(* IEC 61131-3 sources: 2026_Projet_YGO_ExcavatriceDragage/CODE_BACKUP/CODE_20260803_avant_ee4d08b/CODEURS, 7 files *)

(* ---- ST_Encoder_Calib.st ---- *)
(* ═══════════════════════════════════════════════════════════════
   🧲 ST_Encoder_Calib — Calibration & référence codeur (1 par treuil, RETAIN)
   ───────────────────────────────────────────────────────────────
   📄 Doc métier : DOC/AF_Partie-09_Fonction_Encoder_v2.1.md
                   DOC/AF_Partie-03_Contrats_Composants_v2.0.md
   🎛️ Une instance RETAIN par treuil (M1_EncoderCalib / M2_EncoderCalib).
   ═══════════════════════════════════════════════════════════════ *)

TYPE ST_Encoder_Calib :
STRUCT
    HomingRefRaw                  : UDINT;   // Valeur brute figée au dernier homing réussi
    LastKnownRawPos                : UDINT;   // Dernier point brut valide connu (§3.7, continu)
    RestartCoherenceTolerancePts    : UDINT := 1000;  // Tolérance redémarrage (~12% PointsPerRev 8192)
    Homed                          : BOOL;    // TRUE dès qu'un référencement a réussi
    HomingSuspect                  : BOOL;    // TRUE si incohérence détectée au redémarrage (§3.7)
END_STRUCT
END_TYPE

(* ---- FB_Encoder_Abs.st ---- *)
(* ═══════════════════════════════════════════════════════════════
   🧲 FB_Encoder_Abs — Acquisition codeur absolu (accès bus EtherCAT)
   ───────────────────────────────────────────────────────────────
   📄 Doc métier : DOC/AF_Partie-09_Fonction_Encoder_v2.1.md §3/§6
                   DOC/AF_Partie-03_Contrats_Composants_v2.0.md
   🎯 Accès bus EtherCAT, statut esclave, extraction positions brutes
      et séquence de Preset SDO (PresetTriggerCmd := 2).
   🧊 Principe « geler sur doute » (§6) : RawPos/AngleRaw/TurnCount
      conservent leur dernière valeur valide si EncoderAvailable = FALSE.
   ═══════════════════════════════════════════════════════════════ *)

// === DECLARATION (à coller dans la partie déclaration du POU FB_Encoder_Abs) ===

FUNCTION_BLOCK PUBLIC FB_Encoder_Abs
VAR_INPUT
    Enable              : BOOL;        // Standard
    Reset               : BOOL;        // Acquittement défaut (front)
    PowerContactorEngaged     : BOOL;        // Standard
    Mode                : E_Mode;      // Standard (contexte, pas encore exploité ce lot)
    RawPosIn            : UDINT;       // Brut EtherCAT (ex. COD1_PosValue, %ID)
    AlarmsIn            : UINT;        // Brut EtherCAT (ex. COD1_Alarms)
    WarningsIn          : UINT;        // Brut EtherCAT (ex. COD1_Warnings) — informatif seulement
    SlaveOperational    : BOOL;        // FB_Diag_Ethercat — esclave EtherCAT opérationnel
    PointsPerRev        : UDINT := 8192;  // Résolution codeur confirmée (Partie10 §3.3)
    PresetRequest       : BOOL;        // Front — piloté par FB_Encoder_Homing via PRG_02_Encoders
    PresetValue         : UDINT;       // Cible brute — piloté par FB_Encoder_Homing (stub 0 ce lot)
    PresetTimeout       : TIME := T#2s;
    PresetTolerancePts  : UDINT := 10; // Tolérance relecture post-preset
END_VAR
VAR_OUTPUT
    Ready               : BOOL;
    Busy                : BOOL;
    Done                : BOOL;
    Error               : BOOL;
    ErrorId             : WORD;        // bit0: "Défaut communication codeur" - alarme/bus codeur ; bit1: "Erreur référencement (timeout)" - preset refusé/timeout
    State               : E_State;
    StateAtError        : E_State;
    RawPos              : UDINT;       // Position brute — GELÉE si EncoderAvailable=FALSE
    EncoderAvailable    : BOOL;
    AngleRaw            : UINT;        // Informatif maintenance : RawPos MOD PointsPerRev
    TurnCount           : UDINT;       // Informatif maintenance : RawPos / PointsPerRev
    PresetAck           : BOOL;        // Pulse 1 cycle — écriture confirmée
    PresetNak           : BOOL;        // Pulse 1 cycle — écriture refusée/timeout
    PresetTriggerCmd    : WORD;        // → à câbler sur COD_PresettTrigCmd (RxPDO)
    CodeSeqTriggerCmd   : WORD;        // → à câbler sur COD_CodeSeqTrigCmd (RxPDO)
    PresetValueOut      : UDINT;       // → à câbler sur COD_PresetValue (RxPDO)
END_VAR
VAR
    ResetEdge           : R_TRIG;
    ErrorEdge           : R_TRIG;
    PresetReqEdge       : R_TRIG;
    PresetTimer         : TON;
    PresetSeqStep       : INT;         // 0=IDLE, 1=pulse CodeSeq, 2=pulse Trig, 3=attente confirmation
    RawDiff             : DINT;
    PresetTimerVisual   : TON;         // Timer pour laisser le temps de voir l'impulsion (1.5s)
END_VAR

// === IMPLEMENTATION (à coller dans le corps ST du POU FB_Encoder_Abs) ===

// 🛑 1. GATE
IF NOT Enable THEN
    EncoderAvailable := FALSE;
    State := E_State.DISABLED;
    Ready := FALSE; Busy := FALSE; Done := FALSE;
    PresetTriggerCmd := 16#0000; CodeSeqTriggerCmd := 16#0000; PresetValueOut := 0;
    PresetSeqStep := 0;
    PresetTimer(IN := FALSE, PT := PresetTimeout);
    PresetTimerVisual(IN := FALSE, PT := T#500MS);
    RETURN;
END_IF;

Ready := TRUE;
State := E_State.READY;

// 🔑 2. RESET FRONT
ResetEdge(CLK := Reset);

// 🔍 3. DIAGNOSTIC BUS / ALARME
IF (AlarmsIn <> 0) OR NOT SlaveOperational THEN
    ErrorId := ErrorId OR 16#0001;
ELSE
    ErrorId := ErrorId AND 16#FFFE; (* Auto-clearing dès que le bus et l'esclave sont OK *)
END_IF;
EncoderAvailable := (ErrorId AND 16#0001) = 0;

// 📥 4. LECTURE POSITION — GELER SUR DOUTE (Partie10 §6)
// Si EncoderAvailable=FALSE : RawPos/AngleRaw/TurnCount conservent leur dernière valeur (pas de RETURN
// global ici pour ne pas geler aussi la séquence preset/l'état — seule la lecture est gelée).
IF EncoderAvailable THEN
    RawPos := RawPosIn;   // 🔧 2026-07-03 : sens de comptage géré côté codeur (CoE 6000h bit0,
                          // startup parameter CODESYS) — voir Partie10 §3bis. Plus de calcul ici.
    AngleRaw := UDINT_TO_UINT(RawPos MOD PointsPerRev);
    TurnCount := RawPos / PointsPerRev;
END_IF;

// 🔧 5. SÉQUENCE PRESET (écriture bus)
// ✅ Confirmé terrain (2026-07-02) : PresettTrigCmd := 2 déclenche le référencement à
//    PresetValue (valeur de commande, pas un masque de bits — corrige l'hypothèse initiale).
// 🔴 CodeSeqTrigCmd : rôle NON identifié (même par l'utilisateur/terrain) — laissé à 0,
//    PAS piloté tant que sa fonction n'est pas confirmée (fiche technique ou essai dédié).
//    Ne jamais lui donner une valeur arbitraire "au cas où".
PresetReqEdge(CLK := PresetRequest);
PresetAck := FALSE; PresetNak := FALSE; // pulses 1 cycle uniquement
CodeSeqTriggerCmd := 16#0000;           // 🔴 non piloté — rôle inconnu, voir note ci-dessus
CASE PresetSeqStep OF
    0: // IDLE
        PresetTriggerCmd := 0;
        IF PresetReqEdge.Q AND EncoderAvailable THEN
            PresetValueOut := PresetValue;
            PresetSeqStep := 1;
            PresetTimer(IN := TRUE, PT := PresetTimeout);
        END_IF;
    1: // Déclenchement preset (laissé actif pendant 0.5s pour confort visuel en simulation/bus)
        PresetTriggerCmd := 2;   // ✅ Valeur confirmée terrain — référence le codeur à PresetValueOut
        RawDiff := UDINT_TO_DINT(RawPos) - UDINT_TO_DINT(PresetValueOut);
        IF ABS(RawDiff) <= UDINT_TO_DINT(PresetTolerancePts) THEN
            PresetTimer(IN := FALSE, PT := PresetTimeout);
            PresetTimerVisual(IN := TRUE, PT := T#500MS);
            IF PresetTimerVisual.Q THEN
                PresetTriggerCmd := 0;
                PresetAck := TRUE;
                PresetSeqStep := 0;
                PresetTimerVisual(IN := FALSE, PT := T#500MS);
            END_IF;
        ELSIF PresetTimer.Q THEN
            PresetTriggerCmd := 0;
            PresetNak := TRUE;
            ErrorId := ErrorId OR 16#0002;
            PresetSeqStep := 0;
            PresetTimer(IN := FALSE, PT := PresetTimeout);
            PresetTimerVisual(IN := FALSE, PT := T#500MS);
        END_IF;
END_CASE;
IF ResetEdge.Q AND (PresetSeqStep = 0) THEN
    ErrorId := ErrorId AND 16#FFFD;
END_IF;

// 🧾 6. ERROR / STATEATERROR
Error := (ErrorId <> 16#0000);
ErrorEdge(CLK := Error);
IF ErrorEdge.Q THEN
    StateAtError := State;
END_IF;

Busy := (PresetSeqStep <> 0);
Done := PresetAck;

(* ---- FB_Encoder_Homing.st ---- *)
(* ═══════════════════════════════════════════════════════════════
   🎯 FB_Encoder_Homing — Référencement codeur nominal ou unitaire MAINT_N2
   ───────────────────────────────────────────────────────────────
   📄 Doc métier : DOC/AF_Partie-09_Fonction_Encoder_v2.1.md §1/§5/§7bis
                   DOC/AF_Partie-03_Contrats_Composants_v2.0.md
   🎯 Rôle : Gestion du flux de homing nominal (capteur haut + cible paramétrable)
      ou unitaire (MAINT_N2, treuil sélectionné).
   🧮 Calcul du point de calage :
      - PresetValue = centre de la plage multi-tour (marge anti-débordement)
      - HomingRefRaw = PresetValue - round(CfgTopSensorPosM × PointsPerRev / CableM_PerRev)
   🧊 Expose ST_Encoder_Calib en VAR_IN_OUT (RETAIN).
   ═══════════════════════════════════════════════════════════════ *)

// === DECLARATION (à coller dans la partie déclaration du POU FB_Encoder_Homing) ===

FUNCTION_BLOCK PUBLIC FB_Encoder_Homing
VAR_INPUT
    Enable               : BOOL;        // Standard
    Reset                : BOOL;        // Acquittement défaut (front) — bits 0/2/3/4/5 (voir §ErrorId)
    PowerContactorEngaged      : BOOL;        // Standard
    Mode                 : E_Mode;      // MAINT_N1 requis pour le flux nominal
    Home                 : BOOL;        // Demande de référencement (front, bouton IHM UNIQUE)
    UnitaryMode          : BOOL;        // TRUE = flux unitaire à cible libre (MAINT_N2 uniquement)
    WinchSelected        : BOOL;        // TRUE = cette instance est le treuil sélectionné
    CfgHomingTargetM        : REAL;        // Cible libre unitaire, limitée à [-99.0 ; +99.0] m
    BtnConfirmCoherence     : BOOL;        // Front — lève le doute §3.7 (bit9), sans réhoming complet
    TopPositionSensor    : BOOL;        // 🔧 2026-07-02 : capteur position haute UNIQUE, COMMUN aux 2 treuils
                                         // (les 2 câbles hissent ensemble le même ensemble mécanique) — câblé
                                         // IDENTIQUEMENT sur les instances M1 ET M2 (PAS un capteur par treuil),
                                         // voir PRG_MAIN.st
    CfgTopSensorPosM   : REAL := 8.5;   // Cible homing nominal (RETAIN site, voir Partie10 §7bis)
    FwdRevSpeedFeedbackOff : BOOL;      // Retour unique "tous contacteurs sens+vitesse retombés" CE TREUIL — arrêt confirmé
    BrakeFeedback        : BOOL;        // Retour contacteur frein CE TREUIL (TRUE = ouvert/desserré — révocation 2026-08-03)
    RawPos               : UDINT;       // Sortie FB_Encoder_Abs (déjà gelée sur doute)
    EncoderAvailable     : BOOL;        // Sortie FB_Encoder_Abs
    PresetAck            : BOOL;        // Pulse — sortie FB_Encoder_Abs (écriture confirmée)
    PresetNak            : BOOL;        // Pulse — sortie FB_Encoder_Abs (écriture refusée/timeout)
    PointsPerRev         : UDINT := 8192;   // Confirmé fiche technique (Partie10 §3.3)
    MultiTurnRevsMax     : UDINT := 4096;   // Confirmé fiche technique (Partie10 §3.3)
    CableM_PerRev        : REAL := 2.0;     // Confirmé terrain 2026-07-02 (Partie10 §2)
    BypassGlobal         : BOOL := FALSE;   // 🌐 Ignore arrêt confirmé et capteur haut (mise en service)
END_VAR
VAR_OUTPUT
    Ready                : BOOL;
    Busy                 : BOOL;
    Done                 : BOOL;        // Pulse 1 cycle — référencement réussi (miroir PresetAck)
    Error                : BOOL;
    ErrorId              : WORD;        // Voir table de bits en en-tête de fichier / doc §5
    State                : E_State;
    StateAtError         : E_State;
    PresetRequest        : BOOL;        // Pulse → FB_Encoder_Abs.PresetRequest
    PresetValue          : UDINT;       // → FB_Encoder_Abs.PresetValue (= HomingRefTargetNominal)
    Homed                : BOOL;        // RETAIN interne, miroir Calib.Homed
    HomingSuspect        : BOOL;        // RETAIN interne, miroir Calib.HomingSuspect
    HomingRefRaw         : UDINT;       // RETAIN interne, miroir Calib.HomingRefRaw → FB_Encoder_Scale
END_VAR
VAR_IN_OUT
    Calib                : ST_Encoder_Calib;   // Référence vers l'état persistant global (survit aux téléchargements)
END_VAR
VAR
    ResetEdge            : R_TRIG;
    ErrorEdge            : R_TRIG;
    HomeEdge             : R_TRIG;
    ConfirmCoherenceEdge : R_TRIG;
    InitDone             : BOOL;        // Contrôle cohérence §3.7 fait une fois par session Enable
    ArretConfirme        : BOOL;
    PresetValueCalc      : UDINT;       // = HomingRefTargetNominal (constant tant que PointsPerRev/MultiTurnRevsMax fixes)
    TargetPoints         : DINT;        // Écart signé CfgTopSensorPosM → points, figé pendant la séquence
    TargetPositionM      : REAL;        // Cible retenue : nominale ou unitaire
    RawDiffRestart       : DINT;        // Écart |RawPos - LastKnownRawPos| au redémarrage (§3.7)
END_VAR

// === IMPLEMENTATION (à coller dans le corps ST du POU FB_Encoder_Homing) ===

// 🛑 1. GATE — neutralisation ; on continue toutefois d'exposer le dernier état RETAIN connu
// (FB_Encoder_Scale a besoin de HomingRefRaw même si ce FB est désactivé)
IF NOT Enable OR NOT PowerContactorEngaged THEN
    PresetRequest := FALSE;
    PresetValue := 0;
    State := E_State.DISABLED;
    Ready := FALSE; Busy := FALSE; Done := FALSE;
    InitDone := FALSE;   // Force un nouveau contrôle §3.7 à la prochaine activation
    Homed := Calib.Homed;
    HomingSuspect := Calib.HomingSuspect;
    HomingRefRaw := Calib.HomingRefRaw;
    RETURN;
END_IF;

Ready := TRUE;

// 🔑 2. FRONTS
ResetEdge(CLK := Reset);
HomeEdge(CLK := Home);
ConfirmCoherenceEdge(CLK := BtnConfirmCoherence);

// 🔍 3. COHÉRENCE AU REDÉMARRAGE (§3.7) — une fois par session Enable, dès que le codeur répond
IF NOT InitDone THEN
    State := E_State.INIT;
    IF EncoderAvailable THEN
        RawDiffRestart := UDINT_TO_DINT(RawPos) - UDINT_TO_DINT(Calib.LastKnownRawPos);
        IF Calib.Homed AND (ABS(RawDiffRestart) > UDINT_TO_DINT(Calib.RestartCoherenceTolerancePts)) THEN
            Calib.HomingSuspect := TRUE;
            ErrorId := ErrorId OR 16#0200;   // bit9 : incohérence codeur au redémarrage
        END_IF;
        InitDone := TRUE;
    END_IF;
ELSE
    IF State = E_State.INIT THEN State := E_State.READY; END_IF;
END_IF;

// ✅ 4. LEVÉE DU DOUTE (BtnConfirmCoherence, §3.7) — indépendant du Reset générique
IF ConfirmCoherenceEdge.Q AND (Mode = E_Mode.MAINT_N1 OR Mode = E_Mode.MAINT_N2) THEN
    Calib.HomingSuspect := FALSE;
    ErrorId := ErrorId AND 16#FDFF;   // efface bit9
END_IF;

// 🎯 5. DEMANDE DE RÉFÉRENCEMENT (flux nominal)
// Les cibles nominale et unitaire sont rejetées hors du domaine codeur sûr [-99.00;+99.00] m.
// BypassGlobal = TRUE → saute la vérification d'arrêt (mise en service)
ArretConfirme := BypassGlobal OR (FwdRevSpeedFeedbackOff AND NOT BrakeFeedback);

PresetRequest := FALSE;   // Défaut chaque cycle — repose uniquement sur le front HomeEdge ci-dessous
IF HomeEdge.Q AND (State <> E_State.BUSY) THEN
    IF UnitaryMode THEN
        TargetPositionM := CfgHomingTargetM;
    ELSE
        TargetPositionM := CfgTopSensorPosM;
    END_IF;

    // ✅ Homing autorisé en MAINT_N1 et MAINT_N2 — interdit en SEMI_AUTO et en cycle AUTO
    // 🌐 BypassGlobal = TRUE → saute TOUTES les vérifications, force le homing
    IF BypassGlobal THEN
        // Force homing sans condition
        PresetValueCalc := (PointsPerRev * MultiTurnRevsMax) / 2;
        TargetPoints := REAL_TO_DINT(TargetPositionM * UDINT_TO_REAL(PointsPerRev) / CableM_PerRev);
        PresetValue := PresetValueCalc;
        PresetRequest := TRUE;
        State := E_State.BUSY;
    ELSIF (Mode <> E_Mode.MAINT_N1) AND (Mode <> E_Mode.MAINT_N2) THEN
        ErrorId := ErrorId OR 16#0001;        // bit0 : mode non autorisé (seulement MAINT N1/N2)
    ELSIF UnitaryMode AND (Mode <> E_Mode.MAINT_N2) THEN
        ErrorId := ErrorId OR 16#0001;
    ELSIF UnitaryMode AND NOT WinchSelected THEN
        ErrorId := ErrorId OR 16#0002;        // bit1 : mauvais treuil sélectionné
    ELSIF NOT EncoderAvailable THEN
        ErrorId := ErrorId OR 16#0008;        // bit3 : codeur indisponible
    ELSIF NOT ArretConfirme THEN
        ErrorId := ErrorId OR 16#0004;        // bit2 : arrêt non confirmé (contacteurs/frein)
    ELSIF (TargetPositionM < -99.0) OR (TargetPositionM > 99.0) THEN
        ErrorId := ErrorId OR 16#0010;        // bit4 : cible nominale/unitaire hors limites
    ELSIF NOT BypassGlobal AND NOT UnitaryMode AND (TargetPositionM <> 0.0) AND TopPositionSensor THEN
        ErrorId := ErrorId OR 16#0010;        // bit4 : capteur position haute non confirmé
    ELSE
        // ✅ Toutes conditions réunies : calcul de la cible brute et déclenchement
        ErrorId := ErrorId AND 16#FFC0;       // Nettoie les erreurs de rejet 0..5
        PresetValueCalc := (PointsPerRev * MultiTurnRevsMax) / 2;               // Centre exact (§3.3)
        TargetPoints := REAL_TO_DINT(TargetPositionM * UDINT_TO_REAL(PointsPerRev) / CableM_PerRev);
        PresetValue := PresetValueCalc;
        PresetRequest := TRUE;                // Pulse 1 cycle — FB_Encoder_Abs détecte le front lui-même
        State := E_State.BUSY;
    END_IF;
END_IF;

// ⏳ 6. SUIVI DE LA SÉQUENCE (BUSY → confirmation)
Done := FALSE;
IF State = E_State.BUSY THEN
    IF PresetAck THEN
        Calib.HomingRefRaw := DINT_TO_UDINT(UDINT_TO_DINT(PresetValueCalc) - TargetPoints);
        Calib.Homed := TRUE;
        Calib.HomingSuspect := FALSE;
        Calib.LastKnownRawPos := PresetValueCalc;
        Done := TRUE;
        State := E_State.READY;
        // Un homing réussi efface l'intégralité de ErrorId
        ErrorId := 16#0000;
    ELSIF PresetNak THEN
        ErrorId := ErrorId OR 16#0020;        // bit5 : preset refusé/timeout (voir FB_Encoder_Abs)
        State := E_State.READY;
    END_IF;
END_IF;

// 🧾 7. RESET (front) — efface les bits « dernière tentative rejetée » (pas de cause persistante
// à revérifier ici : le prochain Home réévalue toutes les conditions de zéro, voir §5)
IF ResetEdge.Q THEN
    ErrorId := ErrorId AND 16#FFC0;   // efface bits 0..5 (garde bit9, levé seulement par BtnConfirmCoherence/Home)
END_IF;

// 📤 8. SORTIES ÉTAT
Error := (ErrorId <> 16#0000);
ErrorEdge(CLK := Error);
IF ErrorEdge.Q THEN
    StateAtError := State;
END_IF;

// Mise à jour continue du point brut valide connu (hors séquence de homing elle-même)
IF EncoderAvailable AND (State <> E_State.BUSY) THEN
    Calib.LastKnownRawPos := RawPos;
END_IF;

Busy := (State = E_State.BUSY);
Homed := Calib.Homed AND NOT Calib.HomingSuspect; // 🆕 REX 2026-07-08 : Perd l'état homed si suspect (démarrage ou fonctionnement), restauré après BtnConfirmCoherence
HomingSuspect := Calib.HomingSuspect;
HomingRefRaw := Calib.HomingRefRaw;

(* ---- FB_Encoder_Safety.st ---- *)
(* ═══════════════════════════════════════════════════════════════
   🛡️ FB_Encoder_Safety — Bornage physique & relais incohérence redémarrage
   ───────────────────────────────────────────────────────────────
   📄 Doc métier : DOC/AF_Partie-09_Fonction_Encoder_v2.1.md §3.6/§3.7
                   DOC/AF_Partie-03_Contrats_Composants_v2.0.md
   🎯 Rôle :
      - Bornage absolu [-99.00 ; +99.00] m (CablePosMSafe gelée sur dernière valeur plausible).
      - Relais de HomingSuspect (ErrorId bit1).
      - Expose EncoderIncoherent (= Error) consommé par FB_Modes.
   ═══════════════════════════════════════════════════════════════ *)

// === DECLARATION (à coller dans la partie déclaration du POU FB_Encoder_Safety) ===

FUNCTION_BLOCK PUBLIC FB_Encoder_Safety
VAR_INPUT
    Enable           : BOOL;        // Standard
    Reset            : BOOL;        // Acquittement défaut (front) — bit0 uniquement (bit1 suit HomingSuspect, voir §7bis)
    PowerContactorEngaged  : BOOL;        // Standard
    Mode             : E_Mode;      // Standard (contexte, pas encore exploité ce lot)
    CablePosM        : REAL;        // Sortie FB_Encoder_Scale DE CE TREUIL
    HomingSuspect    : BOOL;        // Sortie FB_Encoder_Homing DE CE TREUIL (§3.7, déjà calculé)
    PositionMinM     : REAL := -99.0;  // Bornage physique dur (Partie10 §3.6)
    PositionMaxM     : REAL := 99.0;
    BypassGlobal     : BOOL := FALSE;  // 🌐 Force ErrorId=0, ignore bornage (mise en service)
END_VAR
VAR_OUTPUT
    Ready            : BOOL;
    Busy             : BOOL;
    Done             : BOOL;
    Error            : BOOL;
    ErrorId          : WORD;        // bit0: "Position câble hors plage" - position hors plage physique ; bit1: "Incohérence position boot" - incohérence redémarrage (miroir HomingSuspect)
    State            : E_State;
    StateAtError     : E_State;
    CablePosMSafe    : REAL;        // CablePosM gelée sur dernière valeur plausible si hors plage
    EncoderIncoherent: BOOL;        // = Error — consommé par FB_Modes (refuse SEMI_AUTO)
END_VAR
VAR
    ResetEdge             : R_TRIG;
    ErrorEdge             : R_TRIG;
    LastPlausibleCablePosM: REAL;
END_VAR

// === IMPLEMENTATION (à coller dans le corps ST du POU FB_Encoder_Safety) ===

// 🛑 1. GATE — expose la dernière valeur plausible connue même désactivé
IF NOT Enable THEN
    Ready := FALSE; Busy := FALSE; Done := FALSE;
    State := E_State.DISABLED;
    CablePosMSafe := LastPlausibleCablePosM;
    EncoderIncoherent := FALSE;
    RETURN;
END_IF;

Ready := TRUE;
State := E_State.READY;

// 🔑 2. RESET FRONT
ResetEdge(CLK := Reset);

// 🌐 BYPASS GLOBAL : force ErrorId = 0, ignore bornage et incohérence
IF BypassGlobal THEN
    ErrorId := 16#0000;
END_IF;

// 🔍 3. BORNAGE PHYSIQUE ABSOLU (§3.6) — bit0
IF NOT BypassGlobal AND ((CablePosM < PositionMinM) OR (CablePosM > PositionMaxM)) THEN
    ErrorId := ErrorId OR 16#0001;
ELSE
    ErrorId := ErrorId AND 16#FFFE; (* Auto-clearing dès que la position revient dans la plage valide *)
END_IF;

// 🔍 4. RELAIS INCOHÉRENCE REDÉMARRAGE (§3.7, calculée par FB_Encoder_Homing) — bit1
// Pas d'acquittement ici : la levée se fait via BtnConfirmCoherence/nouveau Home côté
// FB_Encoder_Homing (source), ce FB ne fait QUE relayer l'information pour FB_Modes.
IF NOT BypassGlobal THEN
    IF HomingSuspect THEN
        ErrorId := ErrorId OR 16#0002;
    ELSE
        ErrorId := ErrorId AND 16#FFFD;
    END_IF;
END_IF;

// 🧊 5. GELER SUR DOUTE (§6) — CablePosMSafe ne suit PAS CablePosM si hors plage
IF (ErrorId AND 16#0001) = 16#0000 THEN
    LastPlausibleCablePosM := CablePosM;
END_IF;
CablePosMSafe := LastPlausibleCablePosM;

// 📤 6. SORTIES ÉTAT
Error := (ErrorId <> 16#0000);
ErrorEdge(CLK := Error);
IF ErrorEdge.Q THEN
    StateAtError := State;
END_IF;

EncoderIncoherent := Error;
Busy := FALSE;
Done := FALSE;

(* ---- FB_Encoder_Scale.st ---- *)
(* ═══════════════════════════════════════════════════════════════
   📏 FB_Encoder_Scale — Mise à l'échelle points → mètres (1 par treuil)
   ───────────────────────────────────────────────────────────────
   📄 Doc métier : DOC/AF_Partie-09_Fonction_Encoder_v2.1.md §2/§3.1
                   DOC/AF_Partie-03_Contrats_Composants_v2.0.md
   🎯 Formule : CablePosM = (RawPos - HomingRefRaw) × (CableM_PerRev / PointsPerRev)
   🧮 Arithmétique signée sûre : conversion en DINT avant la soustraction.
   ═══════════════════════════════════════════════════════════════ *)

// === DECLARATION (à coller dans la partie déclaration du POU FB_Encoder_Scale) ===

FUNCTION_BLOCK PUBLIC FB_Encoder_Scale
VAR_INPUT
    RawPos          : UDINT;       // Position brute (sortie FB_Encoder_Abs, déjà gelée sur doute)
    HomingRefRaw    : UDINT;       // Référence brute figée au dernier homing (ST_Encoder_Calib)
    CableM_PerRev   : REAL := 2.0; // Câble déroulé par tour (périmètre tambour confirmé 2026-07-02, réglable site)
    PointsPerRev    : UDINT := 8192; // Résolution codeur confirmée (Partie10 §3.3)
END_VAR
VAR_OUTPUT
    CablePosM       : REAL;        // Position câble en mètres, signée (+ enroulé, − sous l'eau)
END_VAR
VAR
    RawDiff         : DINT;        // Écart signé RawPos - HomingRefRaw (§3.1)
END_VAR

// === IMPLEMENTATION (à coller dans le corps ST du POU FB_Encoder_Scale) ===

// 🧮 Écart signé sûr : conversion DINT AVANT soustraction (§3.1) — jamais l'inverse
RawDiff := UDINT_TO_DINT(RawPos) - UDINT_TO_DINT(HomingRefRaw);

// 📏 Formule fixe points → mètres (Partie10 §2)
IF PointsPerRev > 0 THEN
    CablePosM := DINT_TO_REAL(RawDiff) * (CableM_PerRev / UDINT_TO_REAL(PointsPerRev));
ELSE
    CablePosM := 0.0;   // Garde division par zéro (PointsPerRev mal configuré)
END_IF;

(* ---- FB_Encoder_SpeedMeasure.st ---- *)
(* ═══════════════════════════════════════════════════════════════
   📐 FB_Encoder_SpeedMeasure — Mesure de vitesse câble horodatée
   ───────────────────────────────────────────────────────────────
   📄 Doc : DOC/AF_Partie-09_Fonction_Encoder_v2.1.md §3.8
   🛡️ Sécurité : mesure propriétaire de la chaîne codeur ; aucune réaction machine
   🧩 Dépendances : position sûre fournie par FB_Encoder_Safety
   ═══════════════════════════════════════════════════════════════ *)
FUNCTION_BLOCK PUBLIC FB_Encoder_SpeedMeasure
VAR_INPUT
    Enable        : BOOL; // Autorise l'acquisition
    Reset         : BOOL; // Purge immédiate de l'historique
    Position_M    : REAL; // Position câble sûre en mètres
    PositionValid : BOOL; // TRUE si la chaîne codeur garantit la position
END_VAR
VAR_OUTPUT
    Speed_Mps       : REAL; // Vitesse absolue sur la fenêtre horodatée
    SignedSpeed_Mps : REAL; // Vitesse signée : positive montée, négative descente
    Valid           : BOOL; // TRUE après 6 positions couvrant au moins 50 ms
END_VAR
VAR CONSTANT
    WindowTime   : TIME := T#50MS;
    SamplePeriod : TIME := T#10MS;
    SampleCount  : INT := 6;
END_VAR
VAR
    Positions_M : ARRAY[0..5] OF REAL;
    Timestamps  : ARRAY[0..5] OF TIME;
    CurrentTimestamp : TIME;
    LastTimestamp    : TIME;
    ElapsedSinceSample : TIME;
    WindowElapsed      : TIME;
    CollectedSamples   : INT;
    Index              : INT;
    TimestampInitialized : BOOL;
END_VAR

// ⏱️ Horodatage natif : le calcul utilise le temps réellement écoulé, jamais un cycle supposé.
CurrentTimestamp := TIME();

// Purge des six positions sur rupture de confiance : aucune source antérieure ne peut contaminer la mesure.
IF NOT Enable OR Reset OR NOT PositionValid THEN
    Speed_Mps := 0.0;
    SignedSpeed_Mps := 0.0;
    Valid := FALSE;
    CollectedSamples := 0;
    TimestampInitialized := FALSE;
    RETURN;
END_IF;

// 🕒 Première position de la nouvelle fenêtre.
IF NOT TimestampInitialized THEN
    Positions_M[0] := Position_M;
    Timestamps[0] := CurrentTimestamp;
    LastTimestamp := CurrentTimestamp;
    CollectedSamples := 1;
    TimestampInitialized := TRUE;
    Speed_Mps := 0.0;
    SignedSpeed_Mps := 0.0;
    Valid := FALSE;
    RETURN;
END_IF;

// 🛡️ Rebouclage de TIME détecté localement : purge sans réutiliser le delta aberrant (indépendant de T88).
IF CurrentTimestamp < LastTimestamp THEN
    Positions_M[0] := Position_M;
    Timestamps[0] := CurrentTimestamp;
    LastTimestamp := CurrentTimestamp;
    CollectedSamples := 1;
    Speed_Mps := 0.0;
    SignedSpeed_Mps := 0.0;
    Valid := FALSE;
    RETURN;
END_IF;

ElapsedSinceSample := CurrentTimestamp - LastTimestamp;

// 🛡️ Delta nul : aucune division et aucun doublon d'échantillon.
IF ElapsedSinceSample <= T#0MS THEN
    RETURN;
END_IF;

// 📥 Six positions espacées d'au moins 10 ms donnent cinq intervalles sur la fenêtre interne de 50 ms.
IF ElapsedSinceSample >= SamplePeriod THEN
    LastTimestamp := CurrentTimestamp;

    IF CollectedSamples < SampleCount THEN
        Positions_M[CollectedSamples] := Position_M;
        Timestamps[CollectedSamples] := CurrentTimestamp;
        CollectedSamples := CollectedSamples + 1;
    ELSE
        FOR Index := 0 TO 4 DO
            Positions_M[Index] := Positions_M[Index + 1];
            Timestamps[Index] := Timestamps[Index + 1];
        END_FOR;
        Positions_M[5] := Position_M;
        Timestamps[5] := CurrentTimestamp;
    END_IF;

    IF CollectedSamples = SampleCount THEN
        // 🛡️ Ordre temporel et durée minimale contrôlés avant toute conversion/division.
        IF Timestamps[5] >= Timestamps[0] THEN
            WindowElapsed := Timestamps[5] - Timestamps[0];
            IF WindowElapsed >= WindowTime THEN
                SignedSpeed_Mps := (Positions_M[5] - Positions_M[0])
                                   / (UDINT_TO_REAL(TIME_TO_UDINT(WindowElapsed)) / 1000.0);
                Speed_Mps := ABS(SignedSpeed_Mps);
                Valid := TRUE;
            ELSE
                Speed_Mps := 0.0;
                SignedSpeed_Mps := 0.0;
                Valid := FALSE;
            END_IF;
        ELSE
            Speed_Mps := 0.0;
            SignedSpeed_Mps := 0.0;
            Valid := FALSE;
            CollectedSamples := 0;
            TimestampInitialized := FALSE;
        END_IF;
    END_IF;
END_IF;

(* ---- FB_Encoder_SpeedMonitor.st ---- *)
(* ═══════════════════════════════════════════════════════════════════════════════
   🔍 FB_Encoder_SpeedMonitor — Détection de variation brusque de vitesse câble
   ═══════════════════════════════════════════════════════════════════════════════
   📄 Brique standard de diagnostic — aucun pilotage moteur, aucun SafeStop.
   🎯 Compare deux mesures successives de vitesse linéaire câble en m/s.
   🧩 Le seuil et la durée de confirmation sont fournis par l'appelant :
      aucun réglage métier n'est figé dans cette brique.
   🛡️ Une variation confirmée pose ErrorId bit0. Le défaut reste mémorisé
      jusqu'à disparition de la cause et acquittement par front Reset.
   ═══════════════════════════════════════════════════════════════════════════════
   📄 Docs : DOC/AF_Partie-09_Fonction_Encoder_v2.1.md
*)

FUNCTION_BLOCK PUBLIC FB_Encoder_SpeedMonitor
VAR_INPUT
    Enable                     : BOOL;        // Autorise la surveillance
    Reset                      : BOOL;        // Acquittement par front
    PowerContactorEngaged            : BOOL;        // Contexte sécurité global valide
    Mode                       : E_Mode;      // Contexte de fonctionnement
    SpeedMps                   : REAL;        // Vitesse linéaire absolue mesurée (m/s)
    SpeedVariationThresholdMps : REAL;        // Variation minimale à surveiller (m/s)
    SpeedVariationTimeout      : TIME;        // Durée minimale de confirmation
    SpeedStabilityTimeout      : TIME;        // Durée sans variation avant vitesse stable
END_VAR
VAR_OUTPUT
    Ready                  : BOOL;
    Busy                   : BOOL;
    Done                   : BOOL;
    Error                  : BOOL;
    ErrorId                : WORD;        // bit0 : variation vitesse confirmée
    State                  : E_State;
    StateAtError           : E_State;
    SpeedDeltaMps          : REAL;        // Écart absolu entre deux mesures (m/s)
    SpeedVariationDetected : BOOL;        // Seuil dépassé sur le cycle courant
    SpeedVariationConfirmed: BOOL;        // Seuil dépassé pendant la durée requise
    SpeedStable            : BOOL;        // Vitesse stable pendant SpeedStabilityTimeout
END_VAR
VAR
    ResetEdge          : R_TRIG;
    ErrorEdge          : R_TRIG;
    VariationTimer     : TON;
    StabilityTimer     : TON;
    PreviousSpeedMps   : REAL;
    HasPreviousSpeed   : BOOL;
    VariationActive    : BOOL;
END_VAR

// 🛑 1. GATE — désactivation ou AU non réarmé : aucune alarme persistante.
IF NOT Enable OR NOT PowerContactorEngaged THEN
    Ready := FALSE;
    Busy := FALSE;
    Done := FALSE;
    Error := FALSE;
    ErrorId := 16#0000;
    State := E_State.DISABLED;
    SpeedDeltaMps := 0.0;
    SpeedVariationDetected := FALSE;
    SpeedVariationConfirmed := FALSE;
    SpeedStable := FALSE;
    VariationActive := FALSE;
    HasPreviousSpeed := FALSE;
    VariationTimer(IN := FALSE, PT := SpeedVariationTimeout);
    StabilityTimer(IN := FALSE, PT := SpeedStabilityTimeout);
    RETURN;
END_IF;

Ready := TRUE;
Busy := FALSE;
Done := FALSE;
State := E_State.READY;

// 🔑 2. RESET FRONT — l'acquittement n'efface le défaut que si la cause a disparu.
ResetEdge(CLK := Reset);

// 📏 3. CALCUL DE L'ÉCART DE VITESSE — première mesure utilisée comme référence.
IF NOT HasPreviousSpeed THEN
    PreviousSpeedMps := SpeedMps;
    HasPreviousSpeed := TRUE;
    SpeedDeltaMps := 0.0;
ELSE
    SpeedDeltaMps := ABS(SpeedMps - PreviousSpeedMps);
    PreviousSpeedMps := SpeedMps;
END_IF;

// 🔍 4. DÉTECTION BRUTE + FILTRE TEMPOREL — pas de déclenchement si la durée vaut zéro.
VariationActive := HasPreviousSpeed
                   AND (SpeedVariationThresholdMps >= 0.0)
                   AND (SpeedVariationTimeout > T#0ms)
                   AND (SpeedDeltaMps > SpeedVariationThresholdMps);
SpeedVariationDetected := VariationActive;

VariationTimer(IN := VariationActive, PT := SpeedVariationTimeout);
SpeedVariationConfirmed := VariationTimer.Q;
StabilityTimer(IN := HasPreviousSpeed AND NOT VariationActive AND (SpeedStabilityTimeout > T#0ms), PT := SpeedStabilityTimeout);
SpeedStable := StabilityTimer.Q;

IF SpeedVariationConfirmed THEN
    ErrorId := ErrorId OR 16#0001;
ELSIF ResetEdge.Q AND NOT VariationActive THEN
    ErrorId := ErrorId AND 16#FFFE;
END_IF;

// 📤 5. SORTIES D'ÉTAT — diagnostic standard, aucune commande mouvement.
Error := (ErrorId <> 16#0000);
ErrorEdge(CLK := Error);
IF ErrorEdge.Q THEN
    StateAtError := State;
END_IF;
